Fanuc KAREL source: KT00383.KL

PROGRAM KT00383
%NOLOCKGROUP
VAR
  P1: POSITION
  P2: POSITION
  OUT: BOOLEAN
BEGIN
  OUT = P1 <= P2
END KT00383
